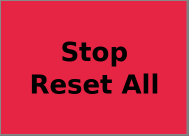
VISUALIZATION OperationButton_Stop  // 189x136
VAR_IN_OUT
	stOperation	:ST_OperationButtons;
END_VAR
    Button (0,0 189x136), "Stop Reset All", colour toggle: stOperation.bStopResetAll, pressed state: stOperation.bStopResetAll
        OnMouseClick: execute { stOperation.bStopResetAll:=TRUE; stOperation.iPauseHistory:=5; }
END_VISUALIZATION

// ---- 00 Library/07-Mode/Visu/Vis_PauseHistory.TcVIS
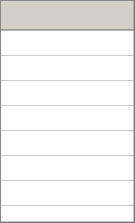
VISUALIZATION Vis_PauseHistory  // 135x223
VAR_IN_OUT
	fbOp: FB_Operation;
END_VAR
    Table (0,0 135x223), data array: fbOp.arPauseHistory
        p3854506369: fbOp.arPauseHistory[INDEX]
        p2232123230: Pause History
END_VISUALIZATION

// ---- 00 Library/10 Utils/DutyCycle/vis_FB_DutyCycle.TcVIS
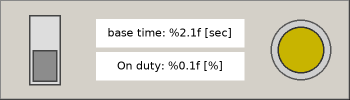
VISUALIZATION vis_FB_DutyCycle  // 350x100
VAR_IN_OUT
	fb: FB_DutyCycle;
END_VAR
    Rectangle (0,0 350x100)
    Lamp1 (266,15 70x70), variable: fb.bOut, style: Lamp-Lamp1-Yellow
    DipSwitch (10,15 70x70), variable: fb.bEnable, behaviour: TOGGLE, style: Switch-DipSwitch-Gray
    Textfield (95,18 150x30), "base time: %2.1f [sec]", text variable: fb.fBaseTime, input disabled if: prg_User.actUser<4
        OnMouseClick: write the text variable via Edit, min 0, max 60
    Textfield (95,51 150x30), "On duty: %0.1f [%]", text variable: fb.fOn_Duty
        OnMouseClick: write the text variable via Edit, min 0, max 100
END_VISUALIZATION

// ---- 00 Library/10 Utils/DutyCycle/vis_FB_DutyCycle_Master.TcVIS
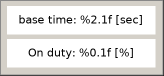
VISUALIZATION vis_FB_DutyCycle_Master  // 164x76
VAR_IN_OUT
	fBaseTime	: REAL;
	fOn_Duty	: REAL;		
END_VAR
    Rectangle (0,0 164x76)
    Textfield (6,5 150x30), "base time: %2.1f [sec]", text variable: fBaseTime
        OnMouseClick: write the text variable via Edit, min 0, max 60
    Textfield (6,38 150x30), "On duty: %0.1f [%]", text variable: fOn_Duty
        OnMouseClick: write the text variable via Edit, min 0, max 100
END_VISUALIZATION

// ---- 01 Instance/04 Recipe/Vis_Recipe_Tab.TcVIS
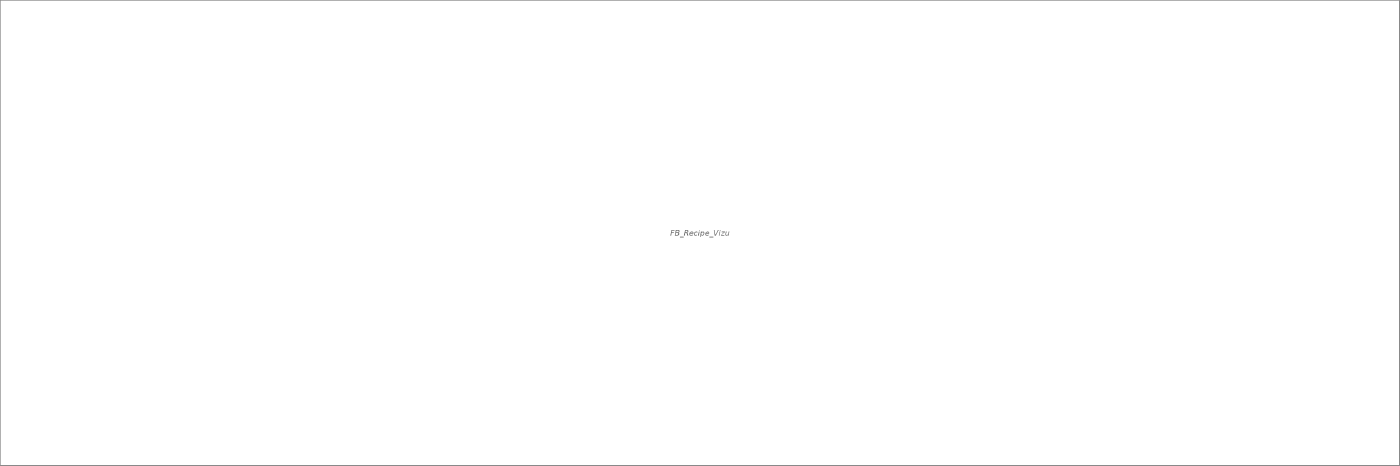
VISUALIZATION Vis_Recipe_Tab  // 1850x617
    TabControl (0,0 1850x617), frame switch variable: prg_Call_Recipe_Slow.iRecipeSwitchFrameVar
        shows FB_Recipe_Vizu(fb_Recipe := GVL_Recipe.fbRecipe[E_Recipe_Name.R_All])
        shows FB_Recipe_Vizu(fb_Recipe := GVL_Recipe.fbRecipe[E_Recipe_Name.R_Device_Dough1])
        shows FB_Recipe_Vizu(fb_Recipe := GVL_Recipe.fbRecipe[E_Recipe_Name.R_Device_Dough2])
        shows FB_Recipe_Vizu(fb_Recipe := GVL_Recipe.fbRecipe[E_Recipe_Name.R_Device_Dough3])
        shows FB_Recipe_Vizu(fb_Recipe := GVL_Recipe.fbRecipe[E_Recipe_Name.R_Device_Dough4])
        shows FB_Recipe_Vizu(fb_Recipe := GVL_Recipe.fbRecipe[E_Recipe_Name.R_CheesyBites])
        shows FB_Recipe_Vizu(fb_Recipe := GVL_Recipe.fbRecipe[E_Recipe_Name.R_CheesyCut])
        shows FB_Recipe_Vizu(fb_Recipe := GVL_Recipe.fbRecipe[E_Recipe_Name.R_Cream])
        shows FB_Recipe_Vizu(fb_Recipe := GVL_Recipe.fbRecipe[E_Recipe_Name.R_Crown])
        shows FB_Recipe_Vizu(fb_Recipe := GVL_Recipe.fbRecipe[E_Recipe_Name.R_Flour])
        shows FB_Recipe_Vizu(fb_Recipe := GVL_Recipe.fbRecipe[E_Recipe_Name.R_Mozzarella])
        shows FB_Recipe_Vizu(fb_Recipe := GVL_Recipe.fbRecipe[E_Recipe_Name.R_Open1])
        shows FB_Recipe_Vizu(fb_Recipe := GVL_Recipe.fbRecipe[E_Recipe_Name.R_Open2])
        shows FB_Recipe_Vizu(fb_Recipe := GVL_Recipe.fbRecipe[E_Recipe_Name.R_Open3])
        shows FB_Recipe_Vizu(fb_Recipe := GVL_Recipe.fbRecipe[E_Recipe_Name.R_Open4])
        shows FB_Recipe_Vizu(fb_Recipe := GVL_Recipe.fbRecipe[E_Recipe_Name.R_Wet])
        shows FB_Recipe_Vizu(fb_Recipe := GVL_Recipe.fbRecipe[E_Recipe_Name.R_Wrap])
        shows FB_Recipe_Vizu(fb_Recipe := GVL_Recipe.fbRecipe[E_Recipe_Name.R_Sesame])
        shows FB_Recipe_Vizu(fb_Recipe := GVL_Recipe.fbRecipe[E_Recipe_Name.R_Piston_Settings])
        [0]: TabTitle=All
        [1]: TabTitle=Device 1
        [2]: TabTitle=Device 2
        [3]: TabTitle=Device 3
        [4]: TabTitle=Device 4
        [5]: TabTitle=Cheesy Bites
        [6]: TabTitle=Cheesy Cut
        [7]: TabTitle=Cream
        [8]: TabTitle=Crown
        [9]: TabTitle=Flour
        [10]: TabTitle=Mozza
        [11]: TabTitle=Open1
        [12]: TabTitle=Open2
        [13]: TabTitle=Open3
        [14]: TabTitle=Open4
        [15]: TabTitle=Wet
        [16]: TabTitle=Wrap
        [17]: TabTitle=Sesame
        [18]: TabTitle=Piston Param
END_VISUALIZATION

// ---- 01 Instance/04-Messages/ERROR_BUFFER.TcVIS
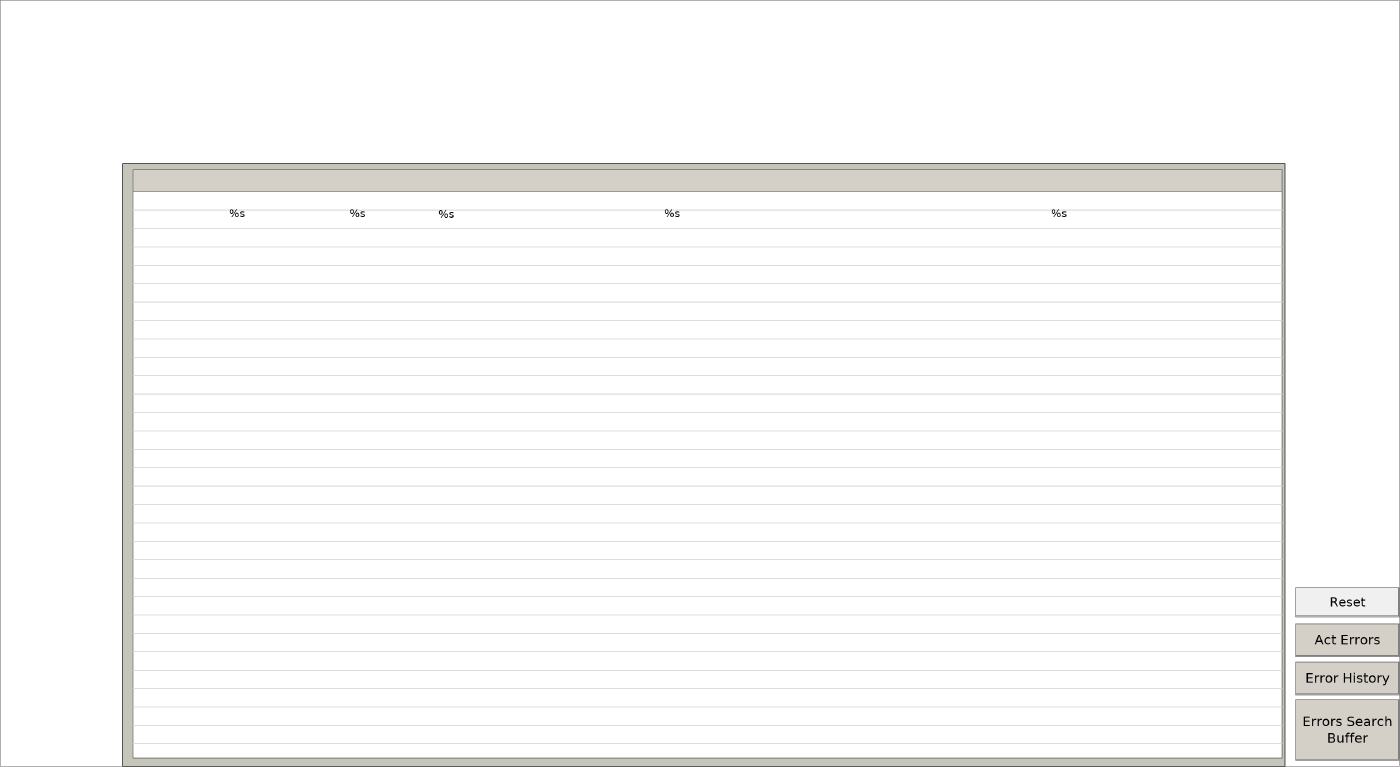
VISUALIZATION ERROR_BUFFER  // 1900x1042
    Group (1758,798 142x235)
        Button (0,0 142x40), "Reset", pressed state: prg_Messages.ResetErrors
            toggle prg_Messages.ResetErrors
        Button (0,101 142x45), "Error History"
            OnMouseClick: change screen: ERROR_HISTORY
        Button (0,152 142x83), "Errors Search Buffer"
            OnMouseClick: change screen: ERROR_BUFFER
        Button (0,49 142x45), "Act Errors"
            OnMouseClick: change screen: ERRORS_OPER
    Rectangle (166,222 1578x820)
    Table (180,230 1560x800), data array: Buffer_Search_Messages
        p3854506369: Buffer_Search_Messages[INDEX].sDateTime
        p1892666644: Buffer_Search_Messages[INDEX].sErrID
        p338671338: Buffer_Search_Messages[INDEX].sLevel
        p2170511999: Buffer_Search_Messages[INDEX].sModuleDescription
        p3723444502: Buffer_Search_Messages[INDEX].sErrorMessage
        p4092479075: Module Description
        p2237128397: Error Message
    Rectangle (421,270 129x40), "%s", text variable: Prg_Filter_Messages.stFilter.sErrID
        OnMouseClick: write the text variable via Edit
    Rectangle (551,271 110x40), "%s", text variable: Prg_Filter_Messages.stFilter.sLevel
        OnMouseClick: write the text variable via Edit
    Rectangle (662,270 501x40), "%s", text variable: Prg_Filter_Messages.stFilter.sModuleDescription
        OnMouseClick: write the text variable via Edit
    Rectangle (1162,270 551x40), "%s", text variable: Prg_Filter_Messages.stFilter.sErrorMessage
        OnMouseClick: write the text variable via Edit
    Rectangle (222,270 200x40), "%s", text variable: Prg_Filter_Messages.stFilter.sDateTime
        OnMouseClick: write the text variable via Edit
END_VISUALIZATION

// ---- 01 Instance/04-Messages/ERROR_HISTORY.TcVIS
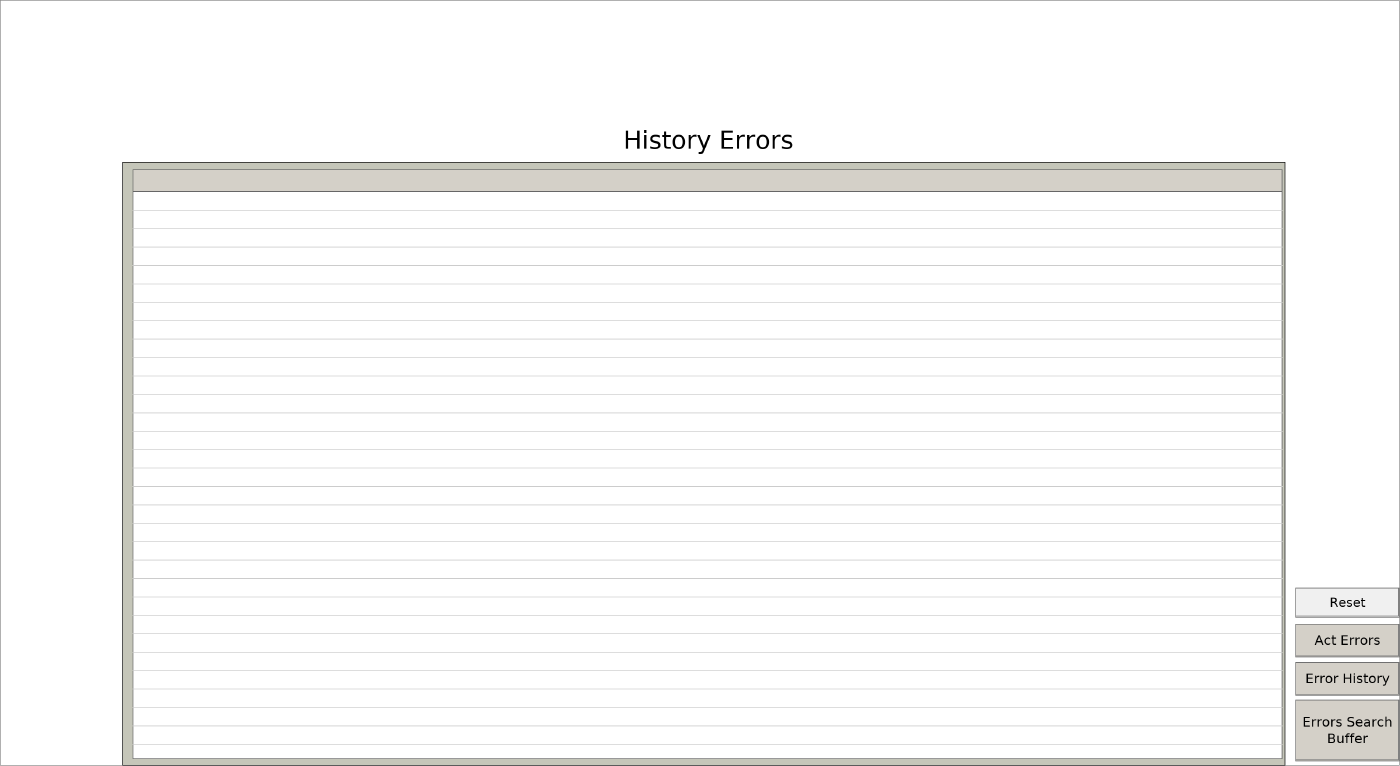
VISUALIZATION ERROR_HISTORY  // 1900x1040
    Group (1758,798 142x235)
        Button (0,0 142x40), "Reset", pressed state: prg_Messages.ResetErrors
            toggle prg_Messages.ResetErrors
        Button (0,101 142x45), "Error History"
            OnMouseClick: change screen: ERROR_HISTORY
        Button (0,152 142x83), "Errors Search Buffer"
            OnMouseClick: change screen: ERROR_BUFFER
        Button (0,49 142x45), "Act Errors"
            OnMouseClick: change screen: ERRORS_OPER
    Rectangle (166,220 1578x820)
    Rectangle (841,165 241x50), "History Errors"
    Table (180,230 1560x800), data array: Buffer_Act_History
        p3854506369: Buffer_Act_History[INDEX].sDateTime
        p1892666644: Buffer_Act_History[INDEX].sErrID
        p338671338: Buffer_Act_History[INDEX].sLevel
        p2170511999: Buffer_Act_History[INDEX].sModuleDescription
        p3723444502: Buffer_Act_History[INDEX].sErrorMessage
        p4092479075: Module Description
        p2237128397: Error Message
END_VISUALIZATION

// ---- 01 Instance/04-Messages/ERROR_Tab.TcVIS
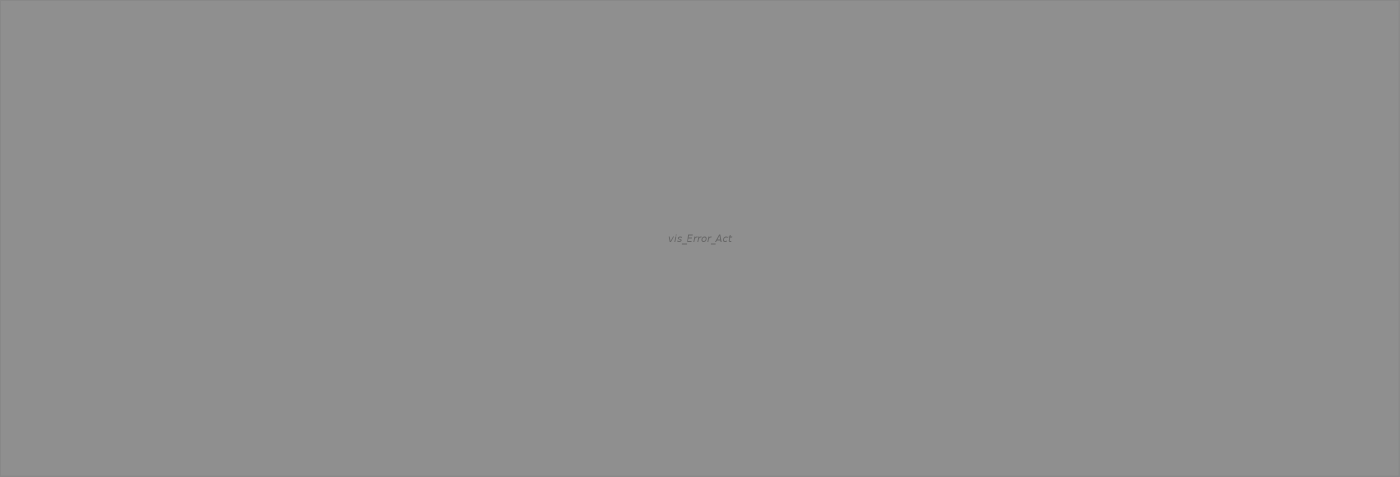
VISUALIZATION ERROR_Tab  // 1428x487
    Rectangle (0,0 1428x487)
    TabControl (0,0 1428x487)
        shows vis_Error_Act()
        shows vis_Error_History()
        shows vis_Error_Search()
        [0]: TabTitle=Actual Errors
        [1]: TabTitle=Error History
        [2]: TabTitle=Search
END_VISUALIZATION

// ---- 01 Instance/04-Messages/ERROR_Tab_1.TcVIS
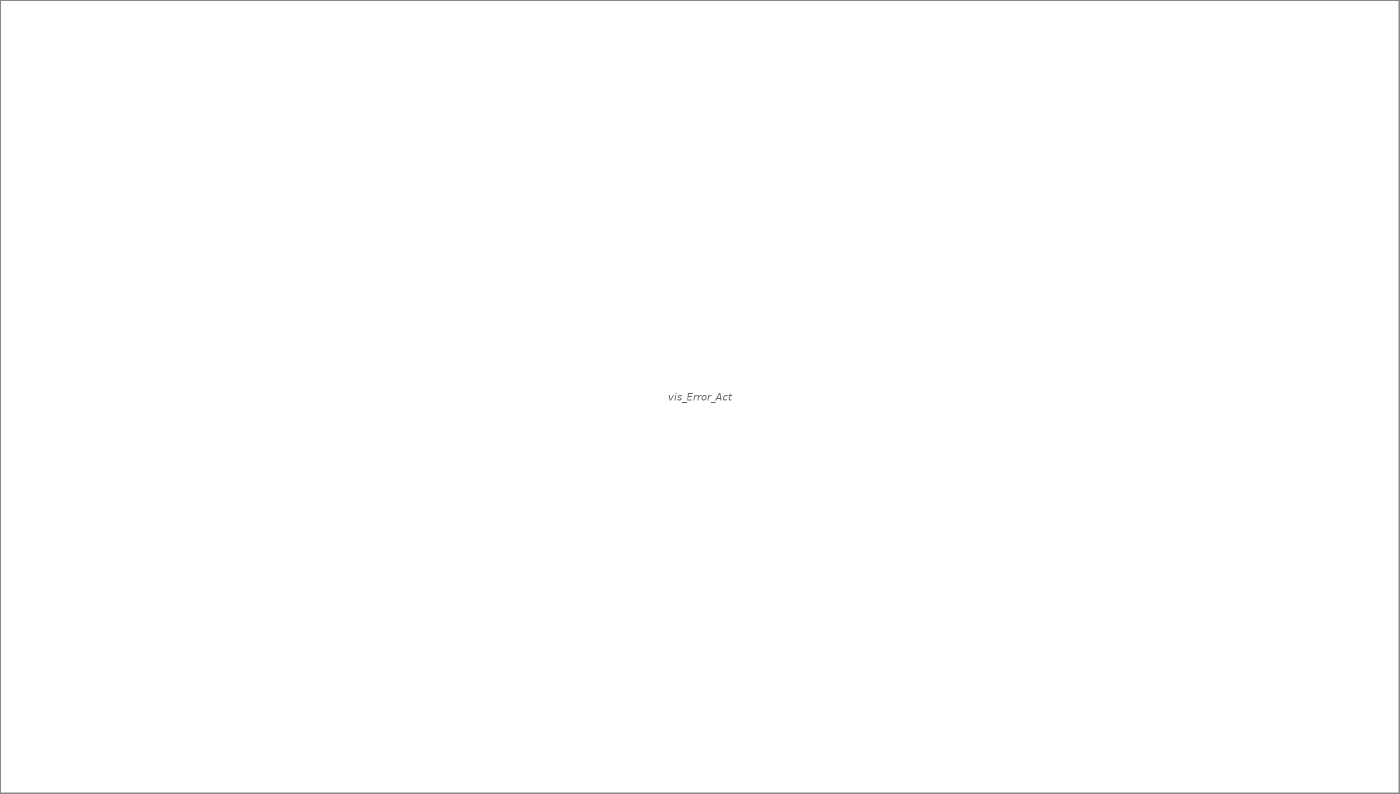
VISUALIZATION ERROR_Tab_1  // 1428x810
    TabControl (0,0 1428x810)
        shows vis_Error_Act()
        shows vis_Error_History()
        shows vis_Error_Search()
        [0]: TabTitle=Actual
        [1]: TabTitle=History
        [2]: TabTitle=Search
END_VISUALIZATION

// ---- 01 Instance/04-Messages/vis_Error_Act.TcVIS
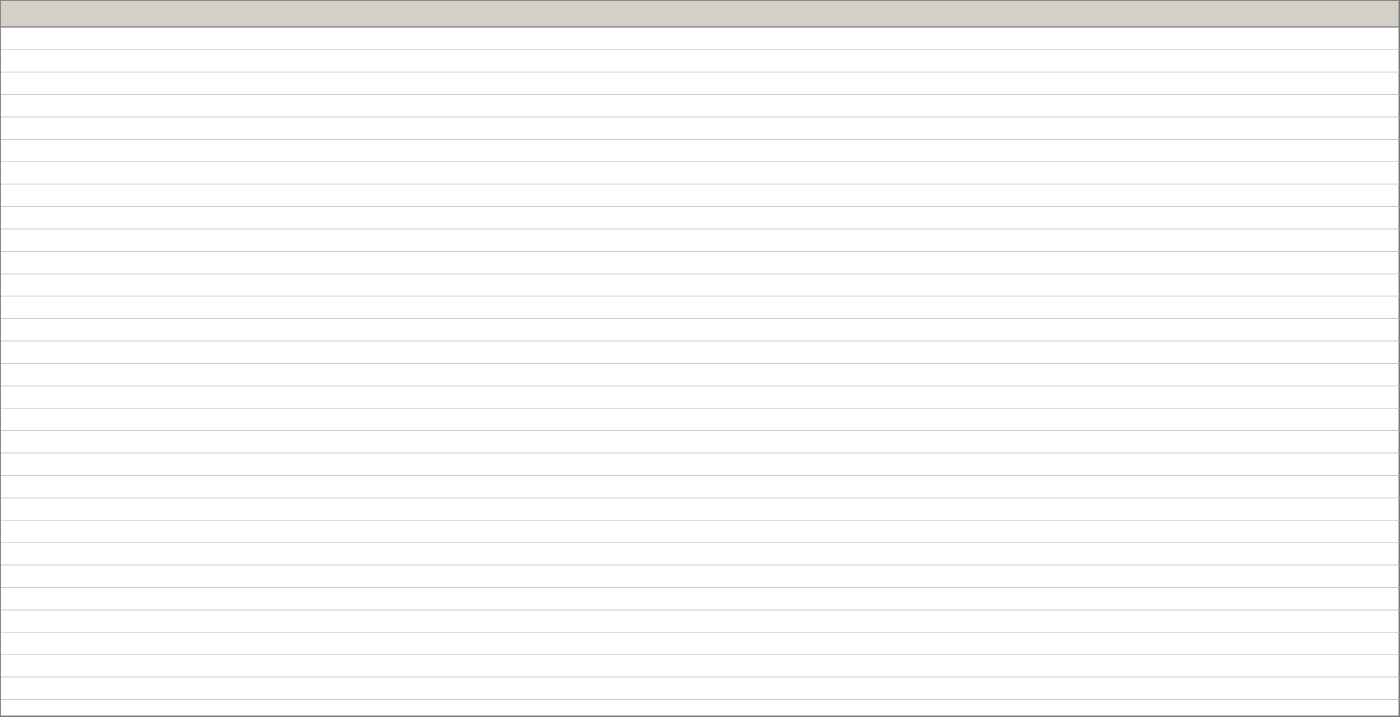
VISUALIZATION vis_Error_Act  // 1560x800
    Table (0,0 1560x800), data array: Buffer_Act_Message
        p3854506369: Buffer_Act_Message[INDEX].sDateTime
        p1892666644: Buffer_Act_Message[INDEX].sErrID
        p338671338: Buffer_Act_Message[INDEX].sLevel
        p2170511999: Buffer_Act_Message[INDEX].sModuleDescription
        p3723444502: Buffer_Act_Message[INDEX].sErrorMessage
        p4092479075: Module Description
        p2237128397: Error Message
END_VISUALIZATION

// ---- 01 Instance/04-Messages/vis_Error_History.TcVIS
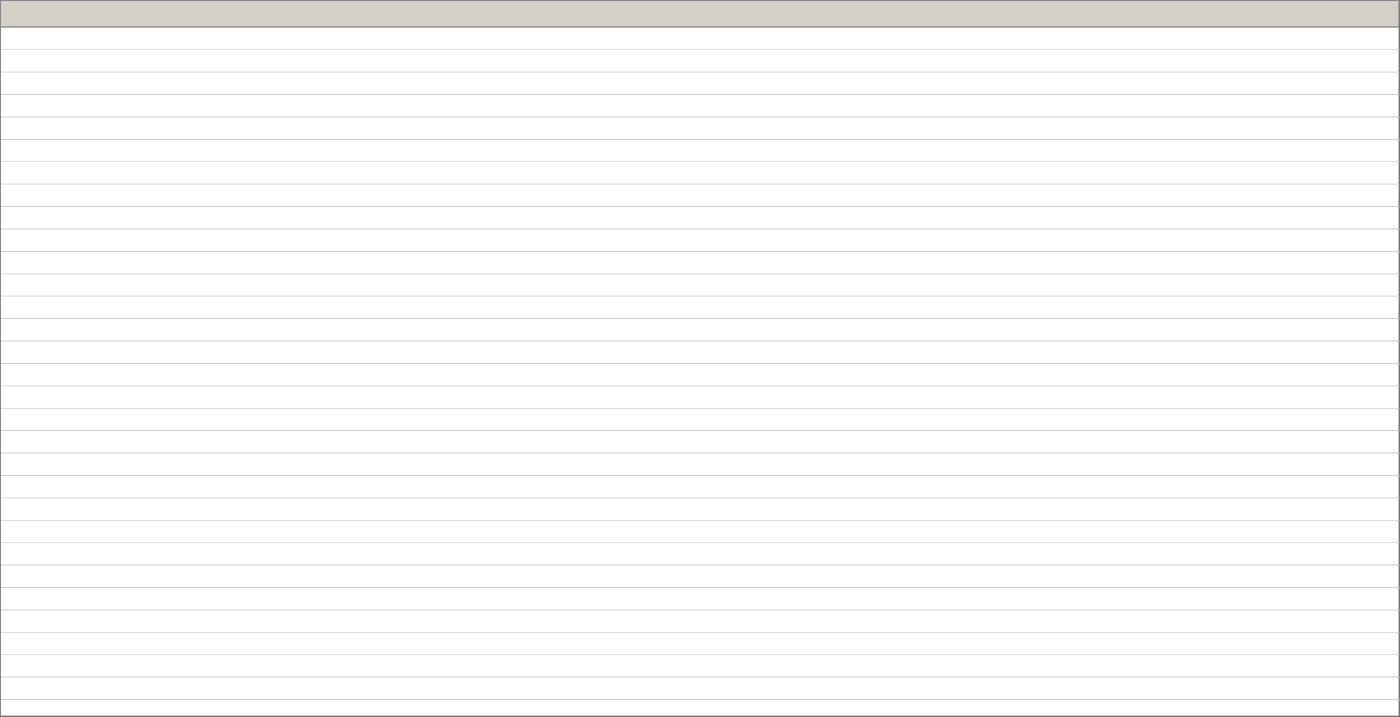
VISUALIZATION vis_Error_History  // 1560x800
    Table (0,0 1560x800), data array: Buffer_Act_History
        p3854506369: Buffer_Act_History[INDEX].sDateTime
        p1892666644: Buffer_Act_History[INDEX].sErrID
        p338671338: Buffer_Act_History[INDEX].sLevel
        p2170511999: Buffer_Act_History[INDEX].sModuleDescription
        p3723444502: Buffer_Act_History[INDEX].sErrorMessage
        p4092479075: Module Description
        p2237128397: Error Message
END_VISUALIZATION

// ---- 01 Instance/04-Messages/vis_Error_Search.TcVIS
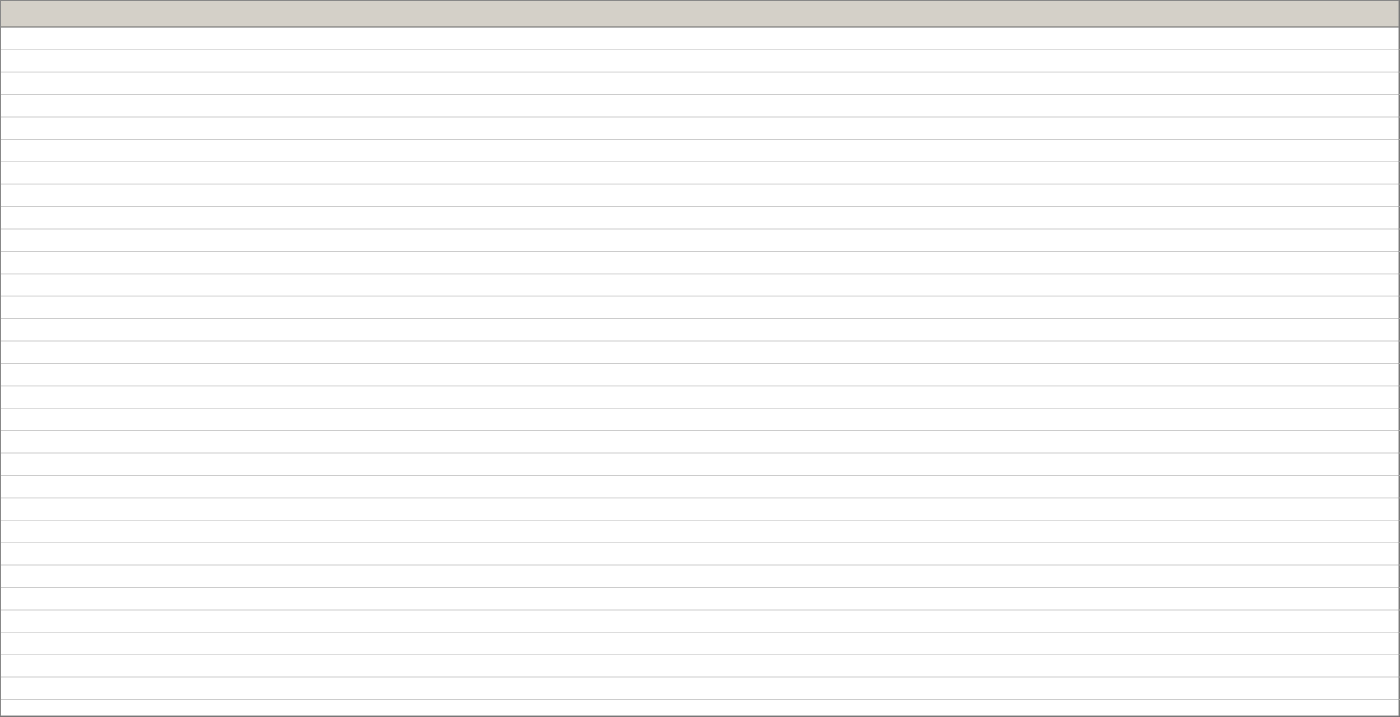
VISUALIZATION vis_Error_Search  // 1560x800
    Table (0,0 1560x800), data array: Buffer_Search_Messages
        p3854506369: Buffer_Search_Messages[INDEX].sDateTime
        p1892666644: Buffer_Search_Messages[INDEX].sErrID
        p338671338: Buffer_Search_Messages[INDEX].sLevel
        p2170511999: Buffer_Search_Messages[INDEX].sModuleDescription
        p3723444502: Buffer_Search_Messages[INDEX].sErrorMessage
        p4092479075: Module Description
        p2237128397: Error Message
END_VISUALIZATION

// ---- 01 Instance/06-Visu/ERRORS_OPER_16_9.TcVIS
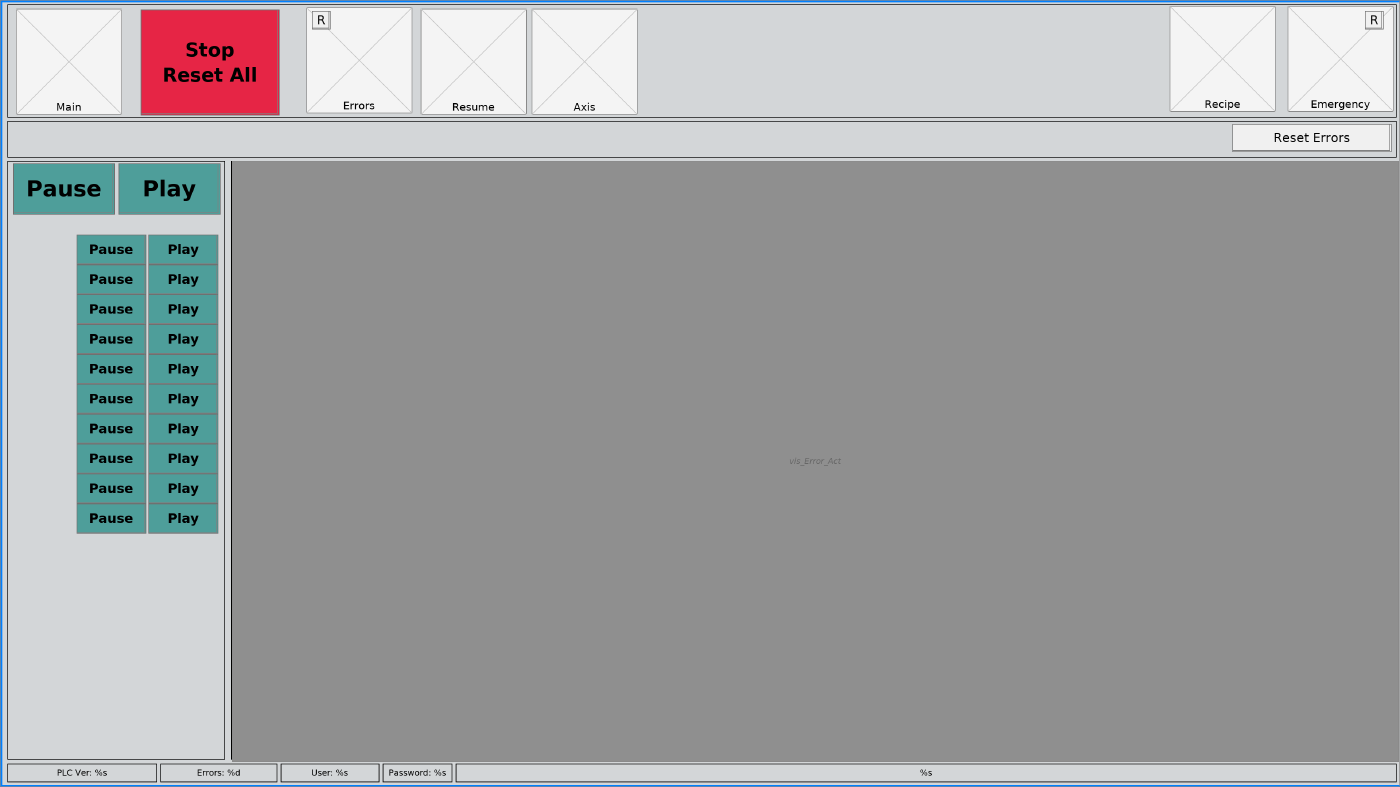
VISUALIZATION ERRORS_OPER_16_9  // 1920x1080
    Frame (0,0 1920x1080)
        shows TEMP16_9_00()
    Frame (318,221 1600x824)
        shows ERROR_Tab()
    Button (1690,170 218x38), "Reset Errors", pressed state: prg_Messages.ResetErrors
        toggle prg_Messages.ResetErrors
END_VISUALIZATION

// ---- 01 Instance/06-Visu/ES_INT_OPER_16_9.TcVIS
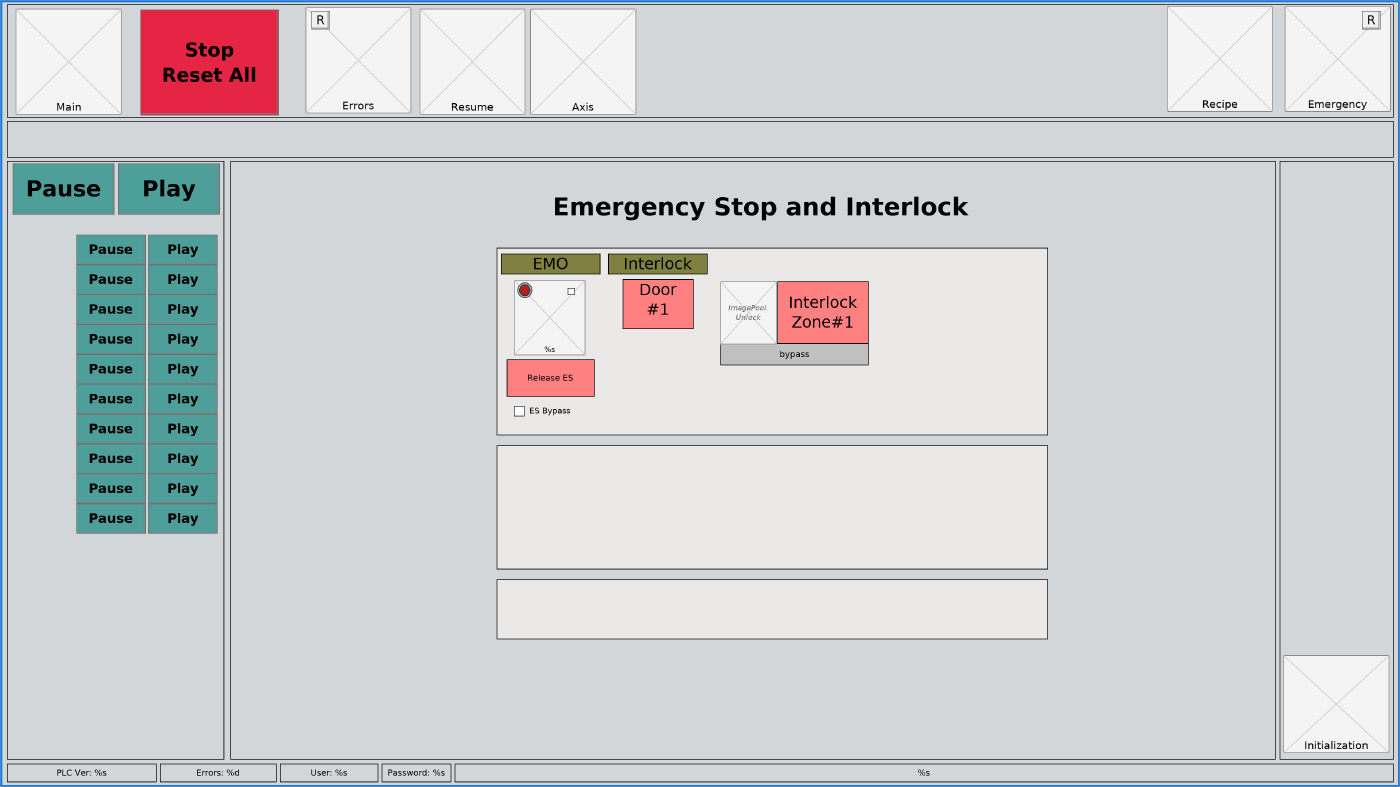
VISUALIZATION ES_INT_OPER_16_9  // 1920x1080
    Frame (0,0 1920x1080)
        shows TEMP16_9_00()
    Rectangle (742,266 602x35), "Emergency Stop and Interlock"
    Rectangle (681,611 756x170)
    Rectangle (681,340 756x257)
    Rectangle (681,795 756x82), invisible if: prg_User.actUser<4
    Rectangle (695,493 120x51), "Release ES", colour toggle: bStateSafe
    Checkbox (703,552 111x24), "ES Bypass", variable: bES_Bypass, invisible if: prg_User.actUser<4
    RoundedRectangle (687,348 136x28), "EMO"
    Frame (705,384 100x103)
        shows Vis_ES_PB(stPB := bES_PB[1], Lable := 'EMO#1')
    RoundedRectangle (834,348 136x28), "Interlock"
    Rectangle (854,383 97x68), "Door #1", colour toggle: bInterlock[1]
    Group (988,386 203x115)
        Rectangle (78,0 125x85), "Interlock Zone#1", colour toggle: bIntZoneLocked[1]
        Rectangle (0,85 203x30), "bypass", colour toggle: bIntZoneBypass[1], invisible if: NOT bIntZoneBypass[1]
            toggle bIntZoneBypass[1]
        Image (0,0 77x86), input disabled if: prg_User.actUser<3, image: ImagePool.Unlock
            p84334746: GVL_Safety.sInterlocksZone1
            OnMouseClick: toggle bIntZoneBypass[1]
END_VISUALIZATION

// ---- 01 Instance/06-Visu/Recipe_16_9.TcVIS
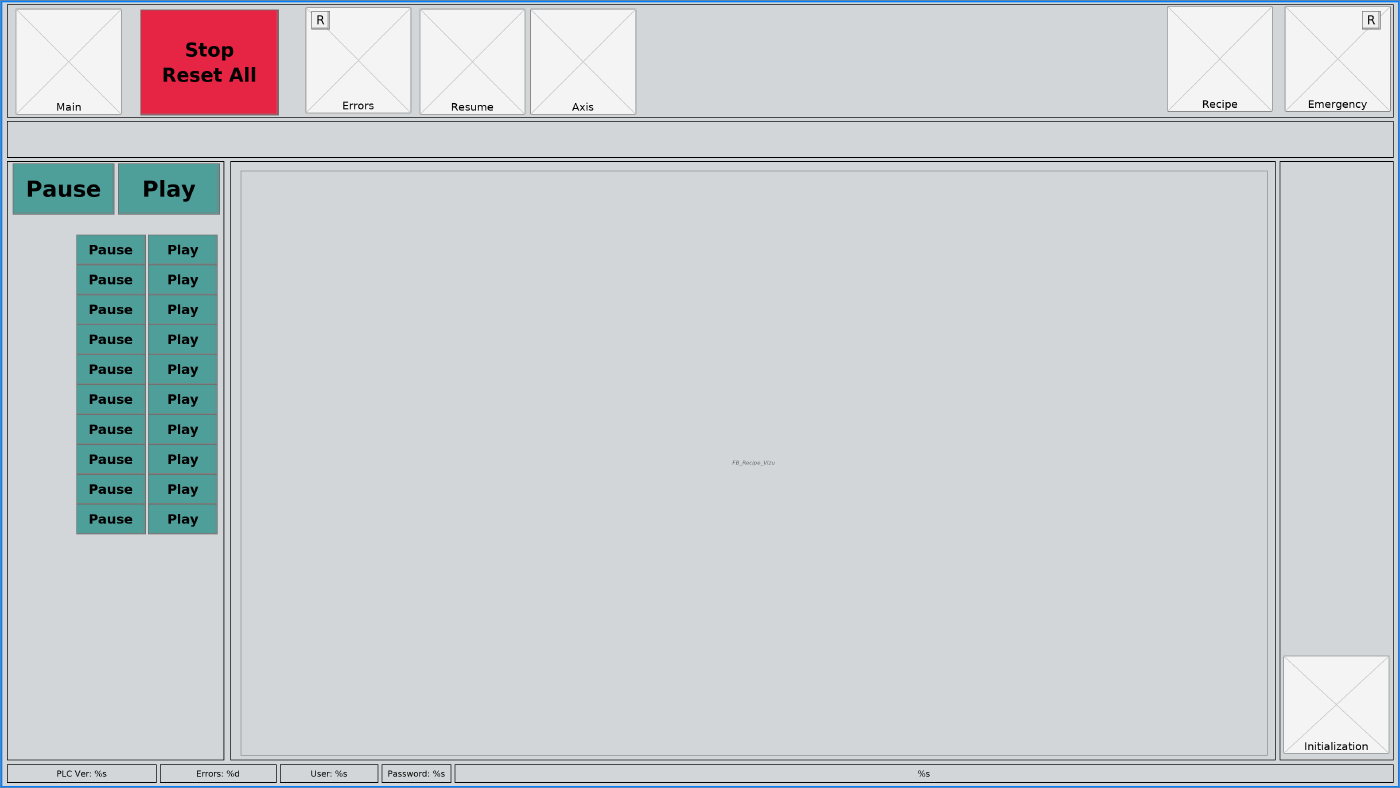
VISUALIZATION Recipe_16_9  // 1920x1081
    Frame (0,0 1920x1081)
        shows TEMP16_9_00()
    Frame (330,234 1408x802)
        shows Vis_Recipe_Tab()
END_VISUALIZATION

// ---- 01 Instance/06-Visu/Template16-9/TEMP16_9_00.TcVIS
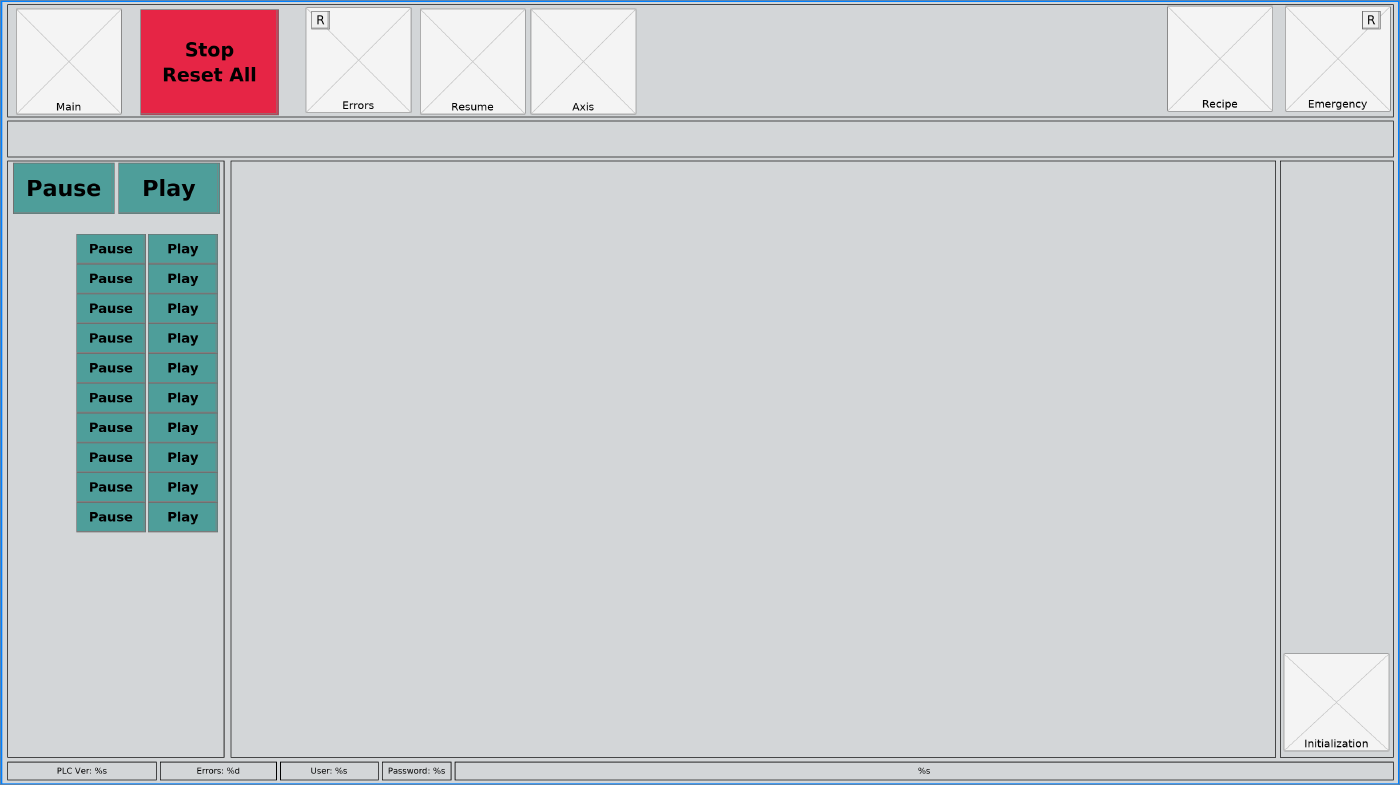
VISUALIZATION TEMP16_9_00  // 1924x1080
    Rectangle (0,0 1924x1080)
    Rectangle (385,1048 135x25), "User: %s", text variable: prg_User.actUser
    Rectangle (525,1048 95x25), "Password: %s", text variable: prg_User.Password
        OnMouseDown: write the text variable via Edit, min 1, max 999
    Rectangle (220,1048 160x25), "Errors: %d", text variable: Global_Persistent.Errors, colour toggle: Global_Persistent.Errors<>0
        OnMouseUp: execute { Global_Persistent.Errors:=(0); }
    Rectangle (10,1048 205x25), "PLC Ver: %s", text variable: ProgramVersion
    Rectangle (625,1048 1290x25), "%s", text variable: sDateTime
    Rectangle (10,6 1905x155)
    Rectangle (10,166 1905x50)
    Image (22,12 145x145), "Main", image: ImagePool.Main
        OnMouseClick: change screen: vis_MAIN
    Image (1766,8 145x145), "Emergency", image: ImagePool.EStop_OK2
        p84334746: GVL_Safety.sBitmap_ESButton
        OnMouseClick: change screen: ES_INT_OPER_16_9
    Image (420,10 145x145), "Errors", image: ImagePool.Error_No
        p84334746: s_Error_BitmapID
        OnMouseClick: change screen: ERRORS_OPER_16_9
    Image (577,12 145x145), "Resume", image: ImagePool.Resume3
        OnMouseClick: toggle ResumeAll
    Button (428,15 25x25), "R", pressed state: prg_Messages.ResetErrors
        toggle prg_Messages.ResetErrors
    Button (1872,15 25x25), "R"
    Rectangle (10,221 298x821)
    Rectangle (1759,221 156x821)
    Frame (18,224 284x70)
        shows OperationButtons(stOperation := stOpMain)
    Image (1764,899 145x134), "Initialization", image: ImagePool.illustration-project-icon
        OnMouseClick: change screen: INIT_OPER_16_9
    Rectangle (317,221 1436x821)
    Frame (193,13 190x145)
        shows OperationButton_Stop(stOperation := stOpMain)
    Image (729,12 145x145), "Axis", image: ImagePool.ervo-motor-beckhoff
        OnMouseClick: change screen: AXIS_OPER
    Image (1604,8 145x145), "Recipe", image: ImagePool.recipe icon
        OnMouseClick: change screen: Recipe_16_9
    Frame (105,322 194x41)
        shows OperationButtons(stOperation := stOper[E_ModeZone.eMain])
    Frame (105,363 194x41)
        shows OperationButtons(stOperation := stOper[E_ModeZone.eCIP])
    Frame (105,404 194x41)
        shows OperationButtons(stOperation := stOper[E_ModeZone.eTank1])
    Frame (105,445 194x41)
        shows OperationButtons(stOperation := stOper[E_ModeZone.eTank2])
    Frame (105,486 194x41)
        shows OperationButtons(stOperation := stOper[E_ModeZone.eTank3])
    Frame (105,527 194x41)
        shows OperationButtons(stOperation := stOper[E_ModeZone.eTank4])
    Frame (105,568 194x41)
        shows OperationButtons(stOperation := stOper[E_ModeZone.eProduction_Marinade])
    Frame (105,609 194x41)
        shows OperationButtons(stOperation := stOper[E_ModeZone.eProduction_Color])
    Frame (105,650 194x41)
        shows OperationButtons(stOperation := stOper[E_ModeZone.eTriBlender_Marinade])
    Frame (105,691 194x41)
        shows OperationButtons(stOperation := stOper[E_ModeZone.eTriBlender_Color])
END_VISUALIZATION

// ---- 01 Instance/06-Visu/Template16-9/TEMP16_9_00_1.TcVIS
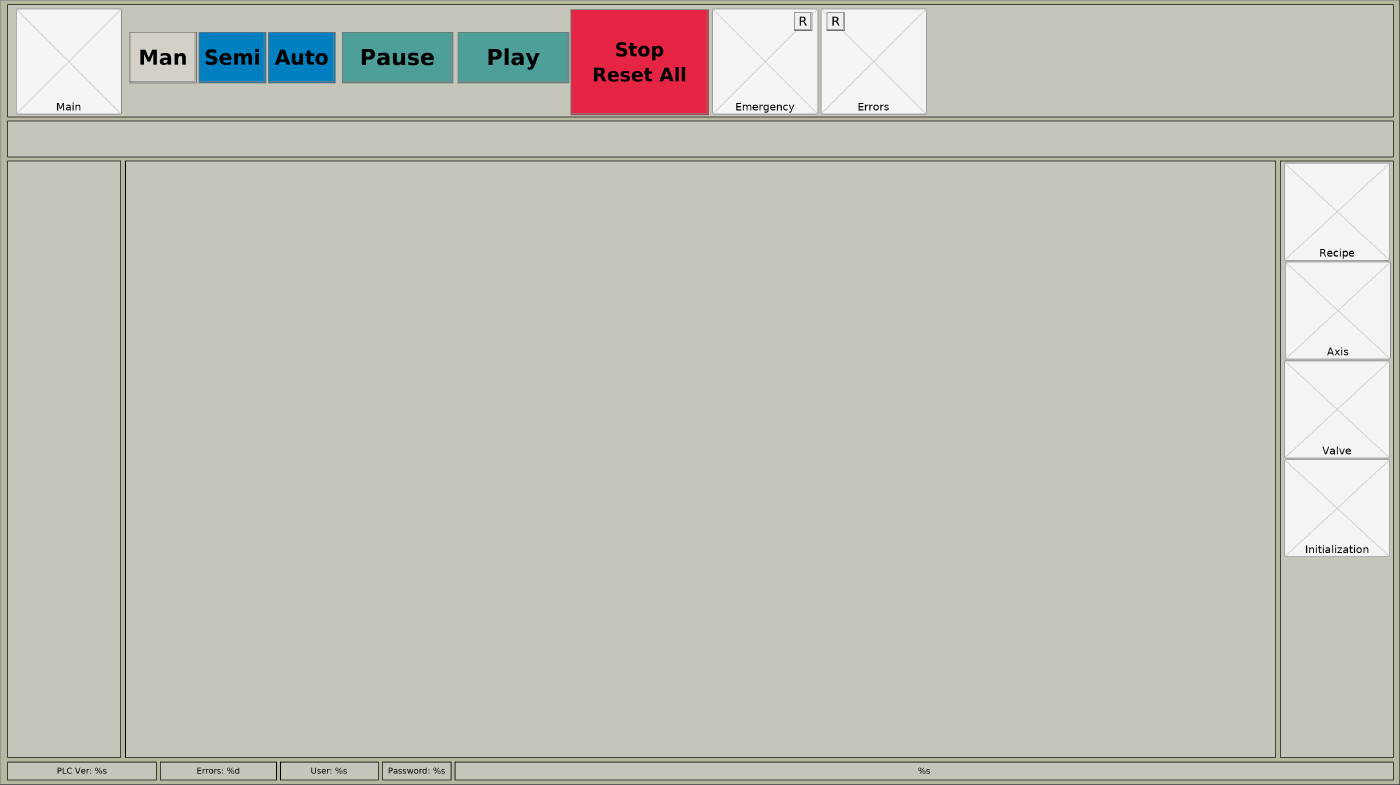
VISUALIZATION TEMP16_9_00_1  // 1924x1080
    Rectangle (0,0 1924x1080)
    Rectangle (385,1048 135x25), "User: %s", text variable: prg_User.actUser
    Rectangle (525,1048 95x25), "Password: %s", text variable: prg_User.Password
        OnMouseDown: write the text variable via Default, min 1, max 999
    Rectangle (220,1048 160x25), "Errors: %d", text variable: Global_Persistent.Errors, colour toggle: Global_Persistent.Errors<>0
        OnMouseUp: execute { Global_Persistent.Errors:=(0); }
    Rectangle (10,1048 205x25), "PLC Ver: %s", text variable: ProgramVersion
    Rectangle (625,1048 1290x25), "%s", text variable: sDateTime
    Rectangle (10,6 1905x155)
    Rectangle (10,166 1905x50)
    Image (22,12 145x145), "Main", image: ImagePool.Main
        OnMouseClick: change screen: vis_MAIN
    Image (979,12 145x145), "Emergency", image: ImagePool.EStop_OK2
        p84334746: GVL_Safety.sBitmap_ESButton
        OnMouseClick: change screen: ES_INT_OPER_16_9
    Image (1128,12 145x145), "Errors", image: ImagePool.Error_No
        p84334746: s_Error_BitmapID
        OnMouseClick: change screen: ERRORS_OPER_16_9
    Button (1136,17 25x25), "R", pressed state: prg_Messages.ResetErrors
        toggle prg_Messages.ResetErrors
    Button (1091,17 25x25), "R"
    Rectangle (10,221 156x821)
    Rectangle (1759,221 156x821)
    Image (1765,224 145x134), "Recipe", image: ImagePool.recipe icon
        OnMouseClick: change screen: Recipe_16_9
    Image (1765,496 145x134), "Valve", image: ImagePool.festo-pistonjpg
        OnMouseClick: change screen: PISTON_OPER_16_9
    Frame (470,44 312x70)
        shows OperationButtons(stOperation := stOpMain)
    Frame (178,44 283x70)
        shows Mode_Select(stMode := stModeMain)
    Image (1765,632 145x134), "Initialization", image: ImagePool.illustration-project-icon
        OnMouseClick: change screen: INIT_OPER_16_9
    Rectangle (172,221 1581x821)
    Frame (784,13 190x145)
        shows OperationButton_Stop(stOperation := stOpMain)
    Image (1766,360 145x134), "Axis", image: ImagePool.ervo-motor-beckhoff
        OnMouseClick: change screen: AXIS_OPER
END_VISUALIZATION

// ---- 01 Instance/06-Visu/Template16-9/TEMP16_9_00_Content.TcVIS
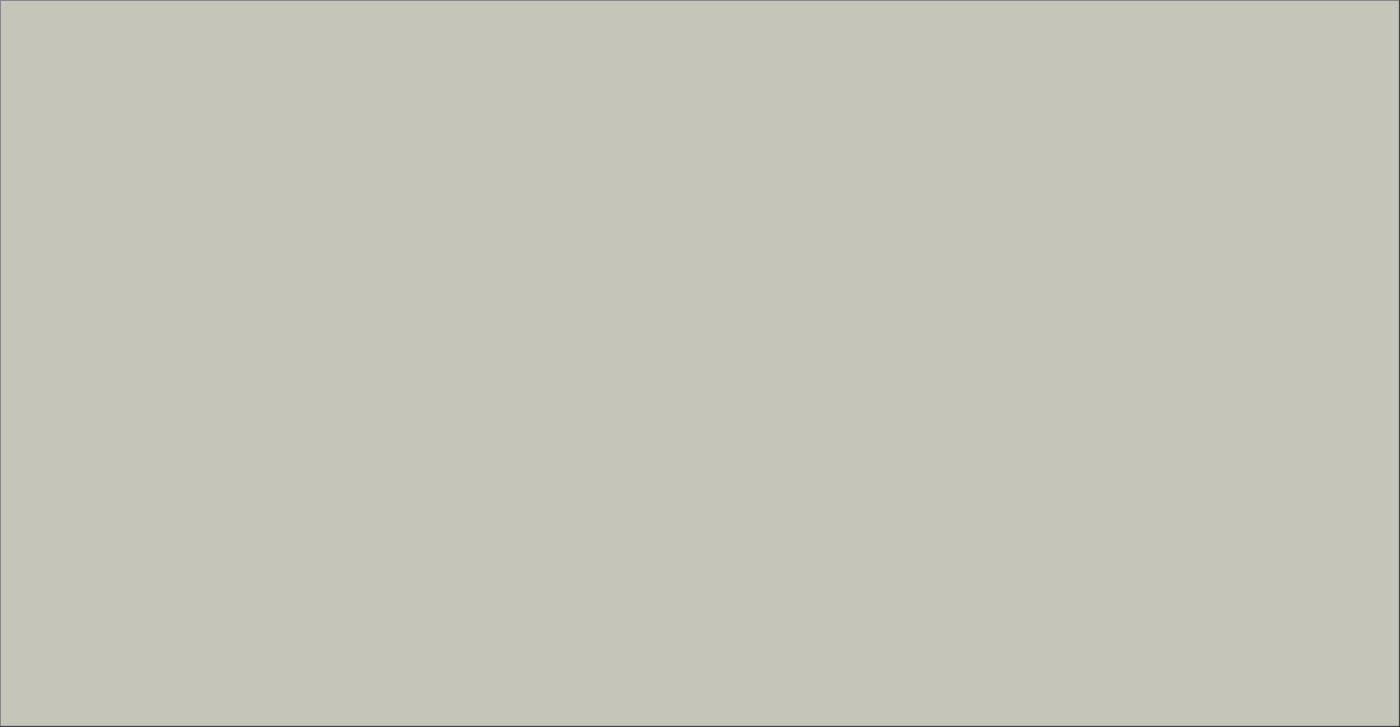
VISUALIZATION TEMP16_9_00_Content  // 1581x821
    Rectangle (0,0 1581x821)
END_VISUALIZATION

// ---- 01 Instance/07-Mode/Vis_LightTower.TcVIS
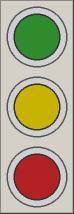
VISUALIZATION Vis_LightTower  // 74x214
    Rectangle (0,0 74x214), colour toggle: prg_LightTower.qBuzzer
    Lamp1 (2,2 70x70), variable: prg_LightTower.qLedGreen, style: Lamp-Lamp1-Green
    Lamp1 (2,72 70x70), variable: prg_LightTower.qLedYellow, style: Lamp-Lamp1-Yellow
    Lamp1 (2,142 70x70), variable: prg_LightTower.qLedRed, style: Lamp-Lamp1-Red
END_VISUALIZATION

// ---- 01 Instance/07-Mode/Vis_LightTower_1.TcVIS
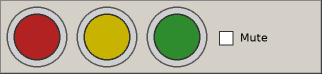
VISUALIZATION Vis_LightTower_1  // 322x74
    Rectangle (0,0 322x74), colour toggle: prg_LightTower.qBuzzer
    Group (2,2 210x70)
        Lamp1 (140,0 70x70), variable: prg_LightTower.qLedGreen, style: Lamp-Lamp1-Green
        Lamp1 (70,0 70x70), variable: prg_LightTower.qLedYellow, style: Lamp-Lamp1-Yellow
        Lamp1 (0,0 70x70), variable: prg_LightTower.qLedRed, style: Lamp-Lamp1-Red
    Checkbox (217,13 95x50), "Mute", variable: bBuzzerMute, input disabled if: prg_User.actUser<2
END_VISUALIZATION

// ---- 01 Instance/07-Mode/viz_HMI_LockIndex.TcVIS
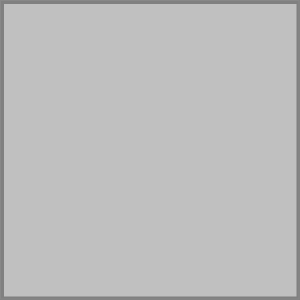
VISUALIZATION viz_HMI_LockIndex  // 300x300
    Rectangle (0,0 300x300), invisible if: not prg_HMI_OperationLock.b_LockIndex
END_VISUALIZATION

// ---- 01 Instance/07-Mode/viz_HMI_Piston.TcVIS
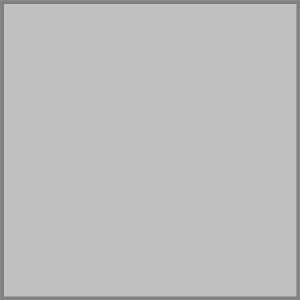
VISUALIZATION viz_HMI_Piston  // 300x300
VAR_INPUT
	bLock_HMI: BOOL;
END_VAR
    Rectangle (0,0 300x300), invisible if: TRUE
END_VISUALIZATION

// ---- 03 Project/23 CIP/TextList_CIP_Clients.TcTLO
TEXTLIST TextList_CIP_Clients
  0 = ' '
  1 = 'Tank1 Marinada'
  2 = 'Tank2 Marinada'
  3 = 'Tank3 Color'
  4 = 'Tank4 Color'
  5 = 'TriBlender Marinada'
  6 = 'TriBlender Color'
  7 = 'Line Marinada'
  8 = 'Line Color'
  9 = 'Local'
   = ''
END_TEXTLIST

// ---- 03 Project/23 CIP/TextList_CIP_Type.TcTLO
TEXTLIST TextList_CIP_Type
  0 = ' '
  1 = 'R Water'
  2 = 'Detergent'
  3 = 'Full'
   = ''
END_TEXTLIST

// ---- 03 Project/23 CIP/vis_CIP.TcVIS
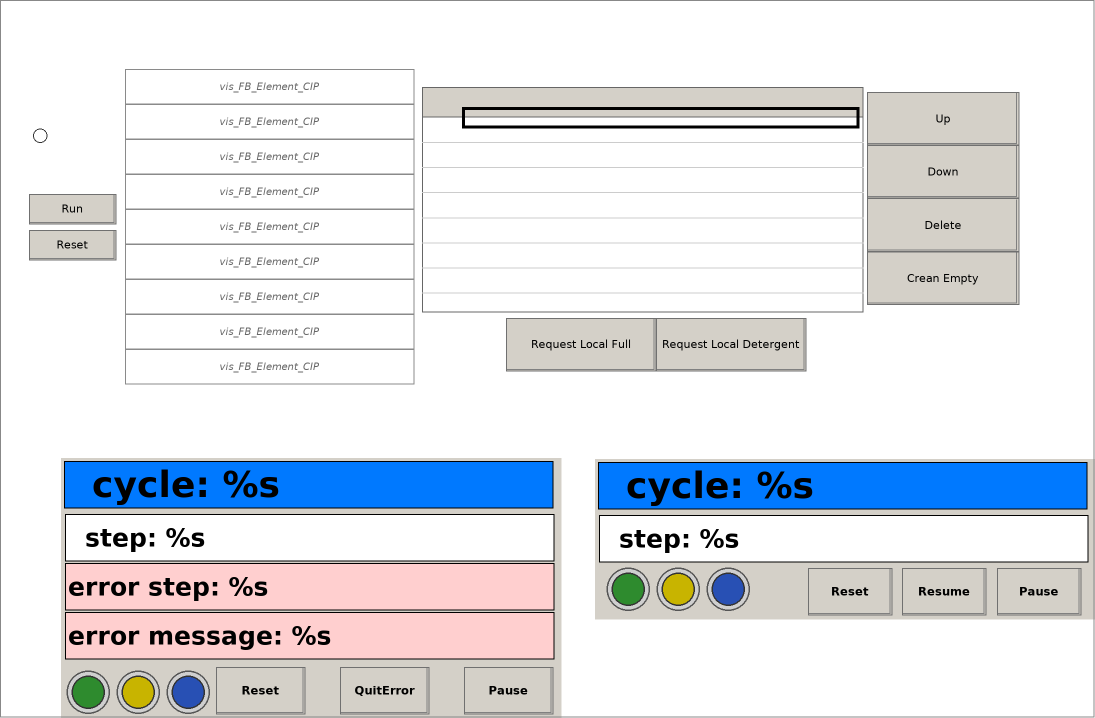
VISUALIZATION vis_CIP  // 1095x718
    Button (29,194 87x30), "Run", colour toggle: fbCIP.bRun
        toggle fbCIP.bRun
    Button (29,230 87x30), "Reset", colour toggle: fbCIP.SFCReset
        toggle fbCIP.SFCReset
    Button (506,318 150x53), "Request Local Full"
        tap fbCIP.rtReqLocalCIP_Full_HMI.CLK
    Button (656,318 150x53), "Request Local Detergent"
        tap fbCIP.rtReqLocalCIP_Detergent_HMI.CLK
    RadioButton (31,86 102x99), variable: fbCIP.eMode
        Areas[0]: Text=Off
        Areas[1]: Text=Manual
        Areas[2]: Text=Auto
    Frame (422,87 597x225)
        shows vis_CIP_ReqBuffer()
    Group (125,69 289x315)
        Frame (0,0 289x35)
            shows vis_FB_Element_CIP(fb := fbElement[E_Element_List.eTank_1])
        Frame (0,35 289x35)
            shows vis_FB_Element_CIP(fb := fbElement[E_Element_List.eTank_2])
        Frame (0,70 289x35)
            shows vis_FB_Element_CIP(fb := fbElement[E_Element_List.eTank_3])
        Frame (0,105 289x35)
            shows vis_FB_Element_CIP(fb := fbElement[E_Element_List.eTank_4])
        Frame (0,140 289x35)
            shows vis_FB_Element_CIP(fb := fbElement[E_Element_List.eTriBlender_Marinada])
        Frame (0,175 289x35)
            shows vis_FB_Element_CIP(fb := fbElement[E_Element_List.eTriBlender_Color])
        Frame (0,210 289x35)
            shows vis_FB_Element_CIP(fb := fbElement[E_Element_List.eLine_Marinada])
        Frame (0,245 289x35)
            shows vis_FB_Element_CIP(fb := fbElement[E_Element_List.eLine_Color])
        Frame (0,280 289x35)
            shows vis_FB_Element_CIP(fb := fbCIP.fbElement_Blank)
    Frame (595,459 500x160)
        shows vis_Cycle_Control(fb := fbCIP, sName := 'CIP')
    Frame (61,458 500x260)
        shows vis_Cycle_Control_1(fb := fbCIP, sName := 'CIP')
END_VISUALIZATION

// ---- 03 Project/23 CIP/vis_CIP_ReqBuffer.TcVIS
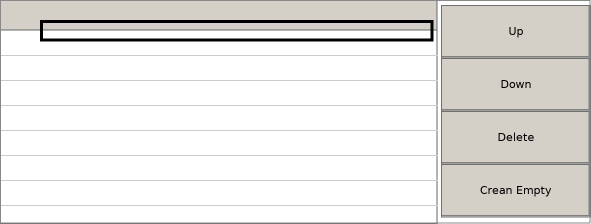
VISUALIZATION vis_CIP_ReqBuffer  // 591x224
    Table (0,0 437x224), data array: arCIP_RequestBufer
        p1137915858: fbCIP.iPosSelect_HMI
        p3854506369: arCIP_RequestBufer[INDEX].eType
        p1892666644: arCIP_RequestBufer[INDEX].eClient
    Button (441,5 150x53), "Up"
        tap fbCIP.rtPosMoveHMI_Up.CLK
    Button (441,58 150x53), "Down"
        tap fbCIP.rtPosMoveHMI_Down.CLK
    Button (441,111 150x53), "Delete"
        tap fbCIP.rtPosDeleteHMI.CLK
    Rectangle (40,20 393x21), colour toggle: fbCIP.bRun
    Button (441,164 150x53), "Crean Empty"
        tap fbCIP.rtReqCleanEmpty_HMI.CLK
END_VISUALIZATION

// ---- 03 Project/31 AnybusCommunication/vis_SiemensSim.TcVIS
